// TIA Portal V21 export
FUNCTION_BLOCK "FB_AnaTimerInner"   // FB17, SCL
TITLE = Analyzer: FB with a timer
{ S7_Optimized_Access := 'TRUE' }
// Rule C26m (callee): the timer is called every time this FB runs
// stored: MemoryReserve 100, SetENOAutomatically false
   VAR_INPUT
      Start : Bool;   // Timer input
   END_VAR
   VAR_OUTPUT
      Done : Bool;   // Timer output
   END_VAR
   VAR
      Delay { S7_SetPoint := 'True'} : TON_TIME;   // On-delay timer
   END_VAR
BEGIN

       #Delay(IN := #Start, PT := T#2s);
       #Done := #Delay.Q;
END_FUNCTION_BLOCK
